FUNCTION_BLOCK Gripper EXTENDS SingleSolenoidCylinder
(*
    Gripper

    A single-solenoid gripper: Extend closes, Retract opens. After the closed
    sensor confirms, the jaws need a moment to build full grip pressure.
*)

PROPERTY PROTECTED SettleTime : TIME
GET
SettleTime := T#150MS;
END_GET
END_PROPERTY

END_FUNCTION_BLOCK

(* stored: Version 1.1.0.1, ProductVersion 3.1.4026.0
   POU Gripper: Id {20dc8eb9-9225-4de5-a77d-3bf4e45ca98b}, SpecialFunc None
   Property SettleTime: Id {c0158ccc-6ed3-45d1-b206-b70b5ceb6cd6}
   Get Get: Id {70fd461b-1a68-43a8-b78c-3401cff58c6c} *)
